(* IEC 61131-3 sources: moqui-plc/codesys-v4/moqui-plc.fbsdev/moqui.iecapp^/moqui/framework/src/start, 2 files *)

(* ---- MoquiStart.prg.st ---- *)
PROGRAM MoquiStart

	VAR
		operationType : OperatingMode := OperatingMode.Init;
		status : MoquiStartStatus := MoquiStartStatus.Idle;
		(* Main framework components *)
		logger : LoggerFacade;
		clockGen : ClockGeneration;
		inputProcessing : InputSignalUpdate;
		outputProcessing : OutputSignalUpdate;
		(* Device config (recipe) management *)
		configMgmt : DeviceConfigMgmt;
		(* Application component *)
		main : Main;
		mainDone : BOOL;
		mainDoneREdge : R_TRIG;
		deviceConfigContextResetRequest : BOOL;
		(*
	     * Keep one Init cycle pending for Main after the first device config has
		 * been loaded, because recipe data also contains device init/homing params.
	     *)
		mainInitPending : BOOL := TRUE;
		(* Error sources: ec.error is written once per cycle from these, so one does not hide the other *)
		configError : BOOL;
		mainError : BOOL;
		(* Reset generated by the retry logic; autoReset belongs to the supervision and is only read here *)
		retryReset : BOOL;
		(* Reset of the device config manager, given on the cycle after a framework reset *)
		configResetRequest : BOOL;
	END_VAR

	(* Set the operating mode *)
	IF ec.init THEN
		(* Logger facade init *)
		logger.enable := TRUE; logger.loggerName := MoquiConf.applicationDeviceId;
		operationType := OperatingMode.Init;
		mainInitPending := TRUE;
	ELSE
		operationType := OperatingMode.Run;
	END_IF;

	(* Timing generation *)
	(*
	 * Uncomment if you want to make loops shorter than 10 ms.
	 * It is not recommended to go below 5 ms with the PLC.
	 * The control loop (current) of the axes is in the servo drives.
	 *)
	(* clks.systemClock := NOT clks.systemClock; *)
	clockGen(operationType := operationType);

	(*
	 * Always run internal procedures, timing generation, process inputs/outputs to ensure safe state
	 * even in software error state, but not in case of hardware/firmware fault.
	 *)
	(* Run hardware fault detection procedures (run network and remote IO diagnostics). *)
	(* runNetworkDgs(error => ec.error);
	IF ec.error THEN
		(* Best if set by an external supervision system: init := FALSE; *)
		status := MoquiStartStatus.Idle;
		RETURN; (* Recycle until the fault condition disappears *)
	END_IF; *)

	(* Input virtualization *)
	(* inputProcessing(operationType := operationType); *)

	(*
	 * Device config (recipe) orchestration must also run during Init because the
	 * first recipe carries the device initialization and homing parameters.
	 *)
	configMgmt(enable := ec.enable, configCompleted := mainDone, reset := configResetRequest,
		allConfigLoaded => ec.allConfigLoaded, error => configError);
	configResetRequest := FALSE;
	(*
	 * Main exposes completion as a level signal; derive a one-scan event here
	 * because recipe advancement and context reset are one-shot actions.
	 *)
	mainDoneREdge(CLK := mainDone);
	IF mainDoneREdge.Q THEN
		deviceConfigContextResetRequest := TRUE;
	END_IF;

	(* Start FMS *)
	CASE status OF
	    MoquiStartStatus.Idle :
			(* Waiting for error reset from supervision *)
	        IF NOT ec.error AND ec.enable THEN
				logger(message := 'Framework started.', level := LogLevel.Info);
	            mainDone := FALSE;
				deviceConfigContextResetRequest := FALSE;
	            status := MoquiStartStatus.Run;
	        END_IF;

	    MoquiStartStatus.Run :
	        IF configMgmt.error THEN
				status := MoquiStartStatus.Error;
	        ELSIF NOT configMgmt.busy THEN
	            IF ec.allConfigLoaded THEN
					logger(message := 'All device configs loaded. Framework idle.', level := LogLevel.Info);
					ec.retryCount := 0; (* A completed run ends the retry sequence *)
					(* Auto disable waiting for new device configs from Moqui or supervision *)
	                ec.enable := FALSE;
	                status := MoquiStartStatus.Idle;
				ELSE
	                (*
	                 * Run the component FSMs sequentially.
					 * The Main component can act as a dispatcher for invoking
	                 * the system's FSM and its subsystems.
					 *
					 * The very first call after recipe load must be Init so that
					 * all device FBs consume their recipe-based init/homing params.
	                 *)
	                main(operationType := SEL(mainInitPending, OperatingMode.Run, OperatingMode.Init),
						enable := ec.enable, deviceConfigContextResetRequest := deviceConfigContextResetRequest,
						done => mainDone, error => mainError);
					mainInitPending := FALSE;
					deviceConfigContextResetRequest := FALSE;
					IF main.error THEN status := MoquiStartStatus.Error; END_IF;
	            END_IF;
	        END_IF;

	    MoquiStartStatus.Error :
	        retryReset := FALSE;
	        (* Retry logic *)
			IF MoquiConf.retryOnError AND (ec.retryCount < MoquiConf.maxRetryCount) THEN
				(* Retry timer update *)
				IF ec.clks.clock1s THEN
					ec.retryTime := ec.retryTime + 1;
				END_IF;

				IF (ec.retryTime >= MoquiConf.minRetryTime) THEN
					logger(message := 'Retrying after error ...', level := LogLevel.Warn);
					ec.retryCount := ec.retryCount + 1;
					ec.retryTime := 0; (* Reset the timer *)
					retryReset := TRUE;
				END_IF;
			END_IF;

	        IF ec.reset OR ec.autoReset OR retryReset THEN
	            logger(message := 'Resetting framework after error.', level := LogLevel.Warn);
	            (* Only a reset from the supervision restarts the retry count: maxRetryCount bounds the automatic ones *)
	            IF ec.reset OR ec.autoReset THEN ec.retryCount := 0; END_IF;
	            retryReset := FALSE;
	            ec.retryTime := 0;
	            mainError := FALSE;
	            configResetRequest := TRUE;
				mainInitPending := TRUE;
				deviceConfigContextResetRequest := FALSE;
	            status := MoquiStartStatus.Idle;
	        END_IF;
	END_CASE;

	(* Single writer of ec.error: the latched Error state, or a device config error still present *)
	ec.error := (status = MoquiStartStatus.Error) OR configError;

	(* Output virtualization *)
	(* outputProcessing(operationType := operationType); *)
	(* Reset the init pulse *)
	ec.init := FALSE;
	END_PROGRAM

(* ---- MqttCommunication.prg.st ---- *)
(*
 * MQTT communication task program: the only caller of the shared connectionFactory.
 *
 * Every cycle it services the broker connection, then the programs that use it, in this order:
 *   1. MqttParameterSub: live parameter writes from Moqui, applied first so that a queued log batch never delays them;
 *   2. MqttParameterPub: optional peer-PLC parameter replication (paramsPubEnable, FALSE by default);
 *   3. LogDispatcher: the log batches (logAppenderEnable).
 * One task owns the MQTT client and all its function blocks, so no other task calls them concurrently.
 *
 * After a connection error the client is disabled, which resets it, and enabled again after mqttReconnectDelay.
 * The connection is opened only while at least one of the three programs is enabled.
 *)
PROGRAM MqttCommunication

	VAR
		connect : BOOL := TRUE;
		reconnectTimer : TON;
		(* Connection errors since start *)
		connectionErrorCount : UDINT;
	END_VAR

	(* An error of the previous cycle disables the client for mqttReconnectDelay *)
	IF connect AND ec.connectionFactory.error THEN
		connect := FALSE;
		IF connectionErrorCount < 16#FFFFFFFF THEN connectionErrorCount := connectionErrorCount + 1; END_IF;
	END_IF;
	reconnectTimer(IN := NOT connect, PT := MoquiConf.mqttReconnectDelay);
	IF reconnectTimer.Q THEN connect := TRUE; END_IF;

	ec.connectionFactory(connect := connect AND (ec.logAppenderEnable OR ec.paramsPubEnable OR ec.paramsSubEnable));

	MqttParameterSub();
	MqttParameterPub();
	LogDispatcher();
	END_PROGRAM
